// Pointeur vers l'axe NC n° nDevice du pool matériel (docs/04 § 6.2) ; 0 si absent
FUNCTION F_AxisRef : POINTER TO AXIS_REF
VAR_INPUT
    nDevice : INT;
END_VAR

IF GVL_IoRef.pAxis = 0 OR nDevice < 1 OR nDevice > GVL_IoRef.nAxes OR nDevice > GVL_Const.MAX_AXES THEN
    F_AxisRef := 0;
ELSE
    F_AxisRef := ADR(GVL_IoRef.pAxis^[nDevice]);
END_IF

END_FUNCTION

(* stored: Version 1.1.0.1, ProductVersion 3.1.4024.12
   POU F_AxisRef: Id {c19fda77-d2e6-535a-940e-9f9a2163bb5a}, SpecialFunc None *)
